// TIA Portal V20 export
// export: Created 2026-10-24T18:20:51.4208089Z, ExportSetting WithDefaults, DisplayName Totally Integrated Automation Portal, DisplayVersion V20 Update 6, DisplayName TIA Portal Openness, DisplayVersion V20 Update 6, DisplayName TIA Portal Version Control Interface, DisplayVersion V20 Update 6, DisplayName SINAMICS Startdrive Advanced, DisplayVersion V20 SP1 Update 2, DisplayName SINAMICS Startdrive G110M, G120, G120C, G120D, G120P, G115D, DisplayVersion V20 SP1 Update 2, DisplayName SINAMICS Startdrive G130, G150, S120, S150, SINAMICS MV, G220, S200, S210, DisplayVersion V20 SP1 Update 2, DisplayName STEP 7 Professional, DisplayVersion V20 Update 6, DisplayName STEP 7 Safety, DisplayVersion V20 Update 2, DisplayName WinCC Basic/Comfort/Advanced, DisplayVersion V20 Update 6, DisplayName WinCC Unified, DisplayVersion V20 Update 6
FUNCTION "FC_FbdLogic" : Void   // FC2, FBD
{ S7_Optimized_Access := 'TRUE' }
VERSION : 0.1
// stored: AutoNumber true, IsIECCheckEnabled false, SetENOAutomatically false, UDAEnableTagReadback false
   VAR_INPUT
      InA : Bool;
      InB : Bool;
   END_VAR
   VAR_OUTPUT
      AndOut : Bool;
      OrOut : Bool;
      XorOut : Bool;
      NotOut : Bool;
      SrOut : Bool;
      RsOut : Bool;
      EdgeOut : Bool;
   END_VAR
   VAR_IN_OUT
      SrBit : Bool;
      RsBit : Bool;
      EdgeBit : Bool;
   END_VAR
   VAR_TEMP   // added for the SCL form of the ladder/FBD networks
      _w1 : Bool;
   END_VAR
BEGIN

REGION Network 1
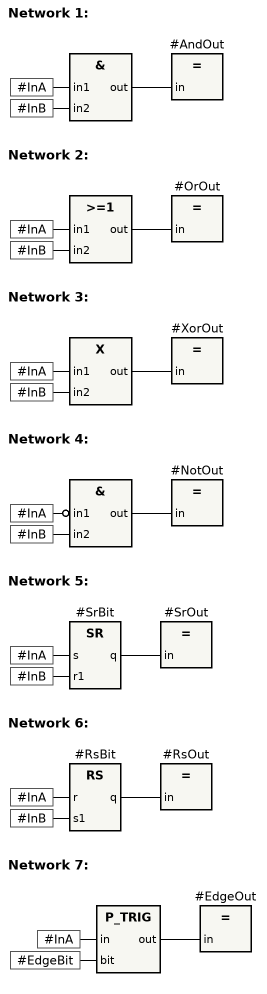
   #AndOut := #InA AND #InB;
END_REGION

REGION Network 2
   #OrOut := #InA OR #InB;
END_REGION

REGION Network 3
   #XorOut := #InA XOR #InB;
END_REGION

REGION Network 4
   #NotOut := NOT #InA AND #InB;
END_REGION

REGION Network 5
   IF #InA THEN
       #SrBit := TRUE;   // SR flip-flop
   END_IF;
   IF #InB THEN #SrBit := FALSE; END_IF;
   #SrOut := #SrBit;
END_REGION

REGION Network 6
   IF #InA THEN
       #RsBit := FALSE;   // RS flip-flop
   END_IF;
   IF #InB THEN #RsBit := TRUE; END_IF;
   #RsOut := #RsBit;
END_REGION

REGION Network 7
   #_w1 := #InA AND NOT #EdgeBit;   // rising edge
   #EdgeBit := #InA;
   #EdgeOut := #_w1;
END_REGION
END_FUNCTION
